              [0]
                bool bANDOR[2]
                num nSigIndex[3]
                num nSigType[3]
                num nValue[3]
            mdesc mMdesc = {leave=0}
            num nActionIndex = 60
            num nDelay = 1
            num nMoveType = 1
            num nPercentage
            num nSigValue = 1
        pointRx pPointRx[2] = {x=-395.706047, y=-287.692007, z=1039.200232, rx=-17.404604, ry=1.457158, rz=-89.580476, shoulder=lefty, elbow=epositive, wrist=wpositive}
        string sID
      [42]
        bool bMarked
        jointRx jJointRx = {j1=-133.481098, j2=-0.271586, j3=94.00243485, j4=-168.691358, j5=107.220034, j6=225.754693}
        pointRx pInter
        paraItem pParaItem
          [0]
            bool bSafePoint
            ifItem iIfItem
              [0]
                bool bANDOR[2]
                num nSigIndex[3]
                num nSigType[3]
                num nValue[3]
            mdesc mMdesc = {leave=0}
            num nActionIndex = 60
            num nDelay = 1
            num nMoveType = 1
            num nPercentage
            num nSigValue = 1
        pointRx pPointRx[2] = {x=-518.840166, y=-287.692002, z=1040.78481, rx=-17.404411, ry=1.457374, rz=-89.580244, shoulder=lefty, elbow=epositive, wrist=wpositive}
        string sID
      [43]
        bool bMarked
        jointRx jJointRx = {j1=-169.544974, j2=-34.564516, j3=135.652231, j4=-196.70666, j5=98.242514, j6=256.952537}
        pointRx pInter
        paraItem pParaItem
          [0]
            bool bSafePoint
            ifItem iIfItem
              [0]
                bool bANDOR[2]
                num nSigIndex[3]
                num nSigType[3]
                num nValue[3]
            mdesc mMdesc = {leave=0}
            num nActionIndex = 60
            num nDelay = 1
            num nMoveType = 1
            num nPercentage
            num nSigValue = 1
        pointRx pPointRx[2] = {x=-445.474256, y=-277.981159, z=882.163294, rx=16.699071, ry=0.613858, rz=-89.857323, shoulder=lefty, elbow=epositive, wrist=wpositive}
        string sID
      [44]
        bool bMarked
        jointRx jJointRx = {j1=-173.644595, j2=-34.491781, j3=138.369342, j4=-179.0487487, j5=104.740151, j6=264.0179677}
        pointRx pInter
        paraItem pParaItem
          [0]
            bool bSafePoint
            ifItem iIfItem
              [0]
                bool bANDOR[2]
                num nSigIndex[3]
                num nSigType[3]
                num nValue[3]
            mdesc mMdesc = {leave=0}
            num nActionIndex = 60
            num nDelay = 1
            num nMoveType = 1
            num nPercentage
            num nSigValue = 1
        pointRx pPointRx[2] = {x=-445.474009, y=-72.78149, z=882.163195, rx=-1.0100742, ry=0.75727, rz=-89.855065, shoulder=lefty, elbow=epositive, wrist=wpositive}
        string sID
      [45]
        bool bMarked
        jointRx jJointRx = {j1=-173.148303, j2=-23.652237, j3=75.107928, j4=-176.801258, j5=42.0835047, j6=260.997576}
        pointRx pInter
        paraItem pParaItem
          [0]
            bool bSafePoint
            ifItem iIfItem
              [0]
                bool bANDOR[2]
                num nSigIndex[3]
                num nSigType[3]
                num nValue[3]
            mdesc mMdesc = {leave=0}
            num nActionIndex = 60
            num nDelay = 1
            num nMoveType = 1
            num nPercentage
            num nSigValue = 1
        pointRx pPointRx[2] = {x=-529.449417, y=-72.791758, z=1365.530984, rx=-1.0242547, ry=-9.601326, rz=-90.0381742, shoulder=lefty, elbow=epositive, wrist=wpositive}
        string sID
      [46]
        bool bMarked
        jointRx jJointRx = {j1=-173.128911, j2=-28.821505, j3=87.506028, j4=-177.167924, j5=49.302114, j6=261.505899}
        pointRx pInter
        paraItem pParaItem
          [0]
            bool bSafePoint
            ifItem iIfItem
              [0]
                bool bANDOR[2]
                num nSigIndex[3]
                num nSigType[3]
                num nValue[3]
            mdesc mMdesc = {leave=0}
            num nActionIndex = 60
            num nDelay = 1
            num nMoveType = 1
            num nPercentage
            num nSigValue = 1
        pointRx pPointRx[2] = {x=-528.694569, y=-72.791769, z=1288.736554, rx=-1.0245197, ry=-9.602488, rz=-90.0383307, shoulder=lefty, elbow=epositive, wrist=wpositive}
        string sID
      [47]
        bool bMarked
        jointRx jJointRx = {j1=-173.184962, j2=-33.03895, j3=99.35319, j4=-177.448656, j5=56.920992, j6=262.0156524}
        pointRx pInter
        paraItem pParaItem
          [0]
            bool bSafePoint
            ifItem iIfItem
              [0]
                bool bANDOR[2]
                num nSigIndex[3]
                num nSigType[3]
                num nValue[3]
            mdesc mMdesc = {leave=0}
            num nActionIndex = 60
            num nDelay = 1
            num nMoveType = 1
            num nPercentage
            num nSigValue = 1
        pointRx pPointRx[2] = {x=-530.992203, y=-72.791768, z=1204.906755, rx=-1.0244931, ry=-9.602628, rz=-90.0383327, shoulder=lefty, elbow=epositive, wrist=wpositive}
        string sID
      [48]
        bool bMarked
        jointRx jJointRx = {j1=-173.214777, j2=-33.556097, j3=101.195834, j4=-177.491533, j5=58.243883, j6=262.117409}
        pointRx pInter
        paraItem pParaItem
          [0]
            bool bSafePoint
            ifItem iIfItem
              [0]
                bool bANDOR[2]
                num nSigIndex[3]
                num nSigType[3]
                num nValue[3]
            mdesc mMdesc = {leave=0}
            num nActionIndex = 60
            num nDelay = 1
            num nMoveType = 1
            num nPercentage
            num nSigValue = 1
        pointRx pPointRx[2] = {x=-532.232127, y=-72.791764, z=1190.718603, rx=-1.0245031, ry=-9.602735, rz=-90.0383446, shoulder=lefty, elbow=epositive, wrist=wpositive}
        string sID
      [49]
        bool bMarked
        jointRx jJointRx = {j1=-170.878262, j2=-41.834096, j3=106.133743, j4=-176.932625, j5=55.0124581, j6=259.371302}
        pointRx pInter
        paraItem pParaItem
          [0]
            bool bSafePoint
            ifItem iIfItem
              [0]
                bool bANDOR[2]
                num nSigIndex[3]
                num nSigType[3]
                num nValue[3]
            mdesc mMdesc = {leave=0}
            num nActionIndex = 60
            num nDelay = 1
            num nMoveType = 1
            num nPercentage
            num nSigValue = 1
        pointRx pPointRx[2] = {x=-459.329518, y=-72.791766, z=1175.87085, rx=-1.0239536, ry=-9.601519, rz=-90.0379744, shoulder=lefty, elbow=epositive, wrist=wpositive}
        string sID
      [50]
        bool bMarked
        jointRx jJointRx = {j1=-164.543315, j2=-49.75207, j3=106.941048, j4=-175.278138, j5=48.290196, j6=251.72242}
        pointRx pInter
        paraItem pParaItem
          [0]
            bool bSafePoint
            ifItem iIfItem
              [0]
                bool bANDOR[2]
                num nSigIndex[3]
                num nSigType[3]
                num nValue[3]
            mdesc mMdesc = {leave=0}
            num nActionIndex = 60
            num nDelay = 1
            num nMoveType = 1
            num nPercentage
            num nSigValue = 1
        pointRx pPointRx[2] = {x=-370.412471, y=-72.791755, z=1185.891907, rx=-1.0250083, ry=-9.601567, rz=-90.0385188, shoulder=lefty, elbow=epositive, wrist=wpositive}
        string sID
      [51]
        bool bMarked
        jointRx jJointRx = {j1=-150.557871, j2=-54.673707, j3=107.498981, j4=-172.114394, j5=45.209263, j6=235.417403}
        pointRx pInter
        paraItem pParaItem
          [0]
            bool bSafePoint
            ifItem iIfItem
              [0]
                bool bANDOR[2]
                num nSigIndex[3]
                num nSigType[3]
                num nValue[3]
            mdesc mMdesc = {leave=0}
            num nActionIndex = 60
            num nDelay = 1
            num nMoveType = 1
            num nPercentage
            num nSigValue = 1
        pointRx pPointRx[2] = {x=-303.196932, y=-72.792593, z=1186.264191, rx=-1.0258078, ry=-9.602273, rz=-90.0389088, shoulder=lefty, elbow=epositive, wrist=wpositive}
        string sID
      [52]
        bool bMarked
        jointRx jJointRx = {j1=-131.882073, j2=-52.891623, j3=101.937702, j4=-168.698385, j5=43.916421, j6=214.126889}
        pointRx pInter
        paraItem pParaItem
          [0]
            bool bSafePoint
            ifItem iIfItem
              [0]
                bool bANDOR[2]
                num nSigIndex[3]
                num nSigType[3]
                num nValue[3]
            mdesc mMdesc = {leave=0}
            num nActionIndex = 60
            num nDelay = 1
            num nMoveType = 1
            num nPercentage
            num nSigValue = 1
        pointRx pPointRx[2] = {x=-265.0832421, y=-72.791017, z=1226.981173, rx=-1.0236731, ry=-9.600494, rz=-90.0378745, shoulder=lefty, elbow=epositive, wrist=wpositive}
        string sID
      [53]
        bool bMarked
        jointRx jJointRx = {j1=-131.398533, j2=-48.129318, j3=93.224241, j4=-167.747499, j5=40.120899, j6=212.404386}
        pointRx pInter
        paraItem pParaItem
          [0]
            bool bSafePoint
            ifItem iIfItem
              [0]
                bool bANDOR[2]
                num nSigIndex[3]
                num nSigType[3]
                num nValue[3]
            mdesc mMdesc = {leave=0}
            num nActionIndex = 60
            num nDelay = 1
            num nMoveType = 1
            num nPercentage
            num nSigValue = 1
        pointRx pPointRx[2] = {x=-264.772643, y=-73.289439, z=1286.811055, rx=-1.0241406, ry=-9.600249, rz=-90.0380209, shoulder=lefty, elbow=epositive, wrist=wpositive}
        string sID
      [54]
        bool bMarked
        jointRx jJointRx = {j1=-144.251884, j2=-41.275682, j3=81.053431, j4=-168.18939, j5=33.105922, j6=224.769818}
        pointRx pInter
        paraItem pParaItem
          [0]
            bool bSafePoint
            ifItem iIfItem
              [0]
                bool bANDOR[2]
                num nSigIndex[3]
                num nSigType[3]
                num nValue[3]
            mdesc mMdesc = {leave=0}
            num nActionIndex = 60
            num nDelay = 1
            num nMoveType = 1
            num nPercentage
            num nSigValue = 1
        pointRx pPointRx[2] = {x=-287.116175, y=-72.447413, z=1363.274189, rx=-1.0263818, ry=-9.602793, rz=-90.03917, shoulder=lefty, elbow=epositive, wrist=wpositive}
        string sID
      [55]
        bool bMarked
        jointRx jJointRx = {j1=-161.427633, j2=-38.278204, j3=80.78039, j4=-172.806947, j5=33.91818, j6=245.804058}
        pointRx pInter
        paraItem pParaItem
          [0]
            bool bSafePoint
            ifItem iIfItem
              [0]
                bool bANDOR[2]
                num nSigIndex[3]
                num nSigType[3]
                num nValue[3]
            mdesc mMdesc = {leave=0}
            num nActionIndex = 60
            num nDelay = 1
            num nMoveType = 1
            num nPercentage
            num nSigValue = 1
        pointRx pPointRx[2] = {x=-347.943507, y=-72.792955, z=1362.805912, rx=-1.0263092, ry=-9.602341, rz=-90.0391422, shoulder=lefty, elbow=epositive, wrist=wpositive}
        string sID
      [56]
        bool bMarked
        jointRx jJointRx = {j1=-168.0500363, j2=-33.981356, j3=79.762569, j4=-175.0248349, j5=36.692248, j6=254.342934}
        pointRx pInter
        paraItem pParaItem
          [0]
            bool bSafePoint
            ifItem iIfItem
              [0]
                bool bANDOR[2]
                num nSigIndex[3]
                num nSigType[3]
                num nValue[3]
            mdesc mMdesc = {leave=0}
            num nActionIndex = 60
            num nDelay = 1
            num nMoveType = 1
            num nPercentage
            num nSigValue = 1
        pointRx pPointRx[2] = {x=-408.635334, y=-72.792697, z=1362.991056, rx=-1.0264229, ry=-9.602398, rz=-90.0392148, shoulder=lefty, elbow=epositive, wrist=wpositive}
        string sID
      [57]
        bool bMarked
        jointRx jJointRx = {j1=-164.68181, j2=-42.542405, j3=92.0793318, j4=-174.620187, j5=40.657851, j6=250.918706}
        pointRx pInter
        paraItem pParaItem
          [0]
            bool bSafePoint
            ifItem iIfItem
              [0]
                bool bANDOR[2]
                num nSigIndex[3]
                num nSigType[3]
                num nValue[3]
            mdesc mMdesc = {leave=0}
            num nActionIndex = 60
            num nDelay = 1
            num nMoveType = 1
            num nPercentage
            num nSigValue = 1
        pointRx pPointRx[2] = {x=-370.383118, y=-72.449044, z=1290.129311, rx=-1.0256153, ry=-9.601833, rz=-90.0387909, shoulder=lefty, elbow=epositive, wrist=wpositive}
        string sID
      [58]
        bool bMarked
        jointRx jJointRx = {j1=-127.503441, j2=-55.600108, j3=106.828006, j4=-168.668567, j5=46.715897, j6=210.0935795}
        pointRx pInter
        paraItem pParaItem
          [0]
            bool bSafePoint
            ifItem iIfItem
              [0]
                bool bANDOR[2]
                num nSigIndex[3]
                num nSigType[3]
                num nValue[3]
            mdesc mMdesc = {leave=0}
            num nActionIndex = 60
            num nDelay = 1
            num nMoveType = 1
            num nPercentage
            num nSigValue = 1
        pointRx pPointRx[2] = {x=-258.489334, y=-72.792581, z=1191.727111, rx=-1.024045, ry=-9.600326, rz=-90.037995, shoulder=lefty, elbow=epositive, wrist=wpositive}
        string sID
      [59]
        bool bMarked
        jointRx jJointRx = {j1=-113.574948, j2=-54.801609, j3=105.785259, j4=-167.709204, j5=48.708352, j6=195.677386}
        pointRx pInter
        paraItem pParaItem
          [0]
            bool bSafePoint
            ifItem iIfItem
              [0]
                bool bANDOR[2]
                num nSigIndex[3]
                num nSigType[3]
                num nValue[3]
            mdesc mMdesc = {leave=0}
            num nActionIndex = 60
            num nDelay = 1
            num nMoveType = 1
            num nPercentage
            num nSigValue = 1
        pointRx pPointRx[2] = {x=-239.513993, y=-72.792586, z=1199.264372, rx=-1.0254298, ry=-9.602381, rz=-90.0386982, shoulder=lefty, elbow=epositive, wrist=wpositive}
        string sID
      [60]
        bool bMarked
        jointRx jJointRx = {j1=-82.821549, j2=-56.0301157, j3=111.780274, j4=-168.953854, j5=58.457299, j6=166.854911}
        pointRx pInter
        paraItem pParaItem
          [0]
            bool bSafePoint
            ifItem iIfItem
              [0]
                bool bANDOR[2]
                num nSigIndex[3]
                num nSigType[3]
                num nValue[3]
            mdesc mMdesc = {leave=0}
            num nActionIndex = 60
            num nDelay = 1
            num nMoveType = 1
            num nPercentage
            num nSigValue = 1
        pointRx pPointRx[2] = {x=-196.990438, y=-72.792703, z=1153.733477, rx=-1.0250656, ry=-9.601957, rz=-90.0385507, shoulder=lefty, elbow=epositive, wrist=wpositive}
        string sID
      [61]
        bool bMarked
        jointRx jJointRx = {j1=-43.782169, j2=-44.715884, j3=104.221439, j4=-173.608416, j5=67.295658, j6=130.959065}
        pointRx pInter
        paraItem pParaItem
          [0]
            bool bSafePoint
            ifItem iIfItem
              [0]
                bool bANDOR[2]
                num nSigIndex[3]
                num nSigType[3]
                num nValue[3]
            mdesc mMdesc = {leave=0}
            num nActionIndex = 60
            num nDelay = 1
            num nMoveType = 1
            num nPercentage
            num nSigValue = 1
        pointRx pPointRx[2] = {x=-98.98037, y=-72.792588, z=1199.212303, rx=-1.0244226, ry=-9.602777, rz=-90.0383225, shoulder=lefty, elbow=epositive, wrist=wpositive}
        string sID
      [62]
        bool bMarked
        jointRx jJointRx = {j1=-33.126092, j2=-38.0272749, j3=100.226244, j4=-175.361365, j5=70.871203, j6=121.320684}
        pointRx pInter
        paraItem pParaItem
          [0]
            bool bSafePoint
            ifItem iIfItem
              [0]
                bool bANDOR[2]
                num nSigIndex[3]
                num nSigType[3]
                num nValue[3]
            mdesc mMdesc = {leave=0}
            num nActionIndex = 60
            num nDelay = 1
            num nMoveType = 1
            num nPercentage
            num nSigValue = 1
        pointRx pPointRx[2] = {x=-39.167207, y=-72.792342, z=1215.189033, rx=-1.0241576, ry=-9.603031, rz=-90.0382398, shoulder=lefty, elbow=epositive, wrist=wpositive}
        string sID
      [63]
        bool bMarked
        jointRx jJointRx = {j1=-26.640244, j2=-32.178556, j3=97.82685, j4=-176.491719, j5=74.724644, j6=115.49475}
        pointRx pInter
        paraItem pParaItem
          [0]
            bool bSafePoint
            ifItem iIfItem
              [0]
                bool bANDOR[2]
                num nSigIndex[3]
                num nSigType[3]
                num nValue[3]
            mdesc mMdesc = {leave=0}
            num nActionIndex = 60
            num nDelay = 1
            num nMoveType = 1
            num nPercentage
            num nSigValue = 1
        pointRx pPointRx[2] = {x=19.131819, y=-72.792471, z=1214.794054, rx=-1.0248151, ry=-9.602165, rz=-90.0383352, shoulder=lefty, elbow=epositive, wrist=wpositive}
        string sID
      [64]
        bool bMarked
        jointRx jJointRx = {j1=-31.251499, j2=-36.639218, j3=99.801437, j4=-180.984741, j5=63.657853, j6=121.825213}
        pointRx pInter
        paraItem pParaItem
          [0]
            bool bSafePoint
            ifItem iIfItem
              [0]
                bool bANDOR[2]
                num nSigIndex[3]
                num nSigType[3]
                num nValue[3]
            mdesc mMdesc = {leave=0}
            num nActionIndex = 60
            num nDelay = 1
            num nMoveType = 1
            num nPercentage
            num nSigValue = 1
        pointRx pPointRx[2] = {x=73.530888, y=-72.792474, z=1249.527518, rx=-1.00980408, ry=0.037023, rz=-89.866745, shoulder=lefty, elbow=epositive, wrist=wpositive}
        string sID
      [65]
        bool bMarked
        jointRx jJointRx = {j1=-29.625602, j2=-33.490872, j3=95.102795, j4=-181.0141949, j5=62.0826287, j6=120.237051}
        pointRx pInter
        paraItem pParaItem
          [0]
            bool bSafePoint
            ifItem iIfItem
              [0]
                bool bANDOR[2]
                num nSigIndex[3]
                num nSigType[3]
                num nValue[3]
            mdesc mMdesc = {leave=0}
            num nActionIndex = 60
            num nDelay = 1
            num nMoveType = 1
            num nPercentage
            num nSigValue = 1
        pointRx pPointRx[2] = {x=89.342541, y=-73.848982, z=1278.496301, rx=-1.00984364, ry=0.0370897, rz=-89.866758, shoulder=lefty, elbow=epositive, wrist=wpositive}
        string sID
      [66]
        bool bMarked
        jointRx jJointRx = {j1=-34.730088, j2=-32.184194, j3=84.304825, j4=-181.0689022, j5=52.670645, j6=125.515286}
        pointRx pInter
        paraItem pParaItem
          [0]
            bool bSafePoint
            ifItem iIfItem
              [0]
                bool bANDOR[2]
                num nSigIndex[3]
                num nSigType[3]
                num nValue[3]
            mdesc mMdesc = {leave=0}
            num nActionIndex = 60
            num nDelay = 1
            num nMoveType = 1
            num nPercentage
            num nSigValue = 1
        pointRx pPointRx[2] = {x=47.85983, y=-72.79225, z=1360.885028, rx=-1.00911117, ry=0.03618, rz=-89.866753, shoulder=lefty, elbow=epositive, wrist=wpositive}
        string sID
      [67]
        bool bMarked
        jointRx jJointRx = {j1=-54.722054, j2=-42.787868, j3=93.663304, j4=-180.780623, j5=51.681236, j6=145.343333}
        pointRx pInter
        paraItem pParaItem
          [0]
            bool bSafePoint
            ifItem iIfItem
              [0]
                bool bANDOR[2]
                num nSigIndex[3]
                num nSigType[3]
                num nValue[3]
            mdesc mMdesc = {leave=0}
            num nActionIndex = 60
            num nDelay = 1
            num nMoveType = 1
            num nPercentage
            num nSigValue = 1
        pointRx pPointRx[2] = {x=-39.660301, y=-72.792082, z=1314.00568418, rx=-1.00941276, ry=0.0361207, rz=-89.866728, shoulder=lefty, elbow=epositive, wrist=wpositive}
        string sID
      [68]
        bool bMarked
        jointRx jJointRx = {j1=-33.267246, j2=-42.513901, j3=112.0835977, j4=-180.919284, j5=70.0957735, j6=123.716984}
        pointRx pInter
        paraItem pParaItem
          [0]
            bool bSafePoint
            ifItem iIfItem
              [0]
                bool bANDOR[2]
                num nSigIndex[3]
                num nSigType[3]
                num nValue[3]
            mdesc mMdesc = {leave=0}
            num nActionIndex = 60
            num nDelay = 1
            num nMoveType = 1
            num nPercentage
            num nSigValue = 1
        pointRx pPointRx[2] = {x=58.0412616, y=-72.792305, z=1160.55849, rx=-1.00998313, ry=0.0362909, rz=-89.866885, shoulder=lefty, elbow=epositive, wrist=wpositive}
        string sID
      [69]
        bool bMarked
        jointRx jJointRx = {j1=-5.272998, j2=-34.693666, j3=109.0300232, j4=-181.0486852, j5=74.39402, j6=95.688496}
        pointRx pInter
        paraItem pParaItem
          [0]
            bool bSafePoint
            ifItem iIfItem
              [0]
                bool bANDOR[2]
                num nSigIndex[3]
                num nSigType[3]
                num nValue[3]
            mdesc mMdesc = {leave=0}
            num nActionIndex = 60
            num nDelay = 1
            num nMoveType = 1
            num nPercentage
            num nSigValue = 1
        pointRx pPointRx[2] = {x=138.724409, y=32.893975, z=1159.616552, rx=-1.010817, ry=0.037884, rz=-89.866801, shoulder=lefty, elbow=epositive, wrist=wpositive}
        string sID
      [70]
        bool bMarked
        jointRx jJointRx = {j1=-4.750773, j2=-30.231867, j3=104.524912, j4=-181.0486754, j5=74.34201, j6=95.167129}
        pointRx pInter
        paraItem pParaItem
          [0]
            bool bSafePoint
            ifItem iIfItem
              [0]
                bool bANDOR[2]
                num nSigIndex[3]
                num nSigType[3]
                num nValue[3]
            mdesc mMdesc = {leave=0}
            num nActionIndex = 60
            num nDelay = 1
            num nMoveType = 1
            num nPercentage
            num nSigValue = 1
        pointRx pPointRx[2] = {x=171.118595, y=32.894004, z=1180.909354, rx=-1.0101343, ry=0.0373213, rz=-89.866785, shoulder=lefty, elbow=epositive, wrist=wpositive}
        string sID
      [71]
        bool bMarked
        jointRx jJointRx = {j1=-4.653989, j2=-28.883061, j3=101.93274, j4=-181.0554282, j5=73.0969745, j6=95.0941538}
        pointRx pInter
        paraItem pParaItem
          [0]
            bool bSafePoint
            ifItem iIfItem
              [0]
                bool bANDOR[2]
                num nSigIndex[3]
                num nSigType[3]
                num nValue[3]
            mdesc mMdesc = {leave=0}
            num nActionIndex = 60
            num nDelay = 1
            num nMoveType = 1
            num nPercentage
            num nSigValue = 1
        pointRx pPointRx[2] = {x=177.941891, y=32.894009, z=1198.169889, rx=-1.0101153, ry=0.0374946, rz=-89.866798, shoulder=lefty, elbow=epositive, wrist=wpositive}
        string sID
      [72]
        bool bMarked
        jointRx jJointRx = {j1=-6.324297, j2=-43.288006, j3=121.304095, j4=-181.0301689, j5=78.0921301, j6=96.670438}
        pointRx pInter
        paraItem pParaItem
          [0]
            bool bSafePoint
            ifItem iIfItem
              [0]
                bool bANDOR[2]
                num nSigIndex[3]
                num nSigType[3]
                num nValue[3]
            mdesc mMdesc = {leave=0}
            num nActionIndex = 60
            num nDelay = 1
            num nMoveType = 1
            num nPercentage
            num nSigValue = 1
        pointRx pPointRx[2] = {x=89.587288, y=32.894025, z=1078.175922, rx=-1.0100336, ry=0.0373229, rz=-89.866767, shoulder=lefty, elbow=epositive, wrist=wpositive}
        string sID
      [73]
        bool bMarked
        jointRx jJointRx = {j1=-29.152055, j2=-40.808391, j3=117.784866, j4=-180.923594, j5=77.436909, j6=119.489453}
        pointRx pInter
        paraItem pParaItem
          [0]
            bool bSafePoint
            ifItem iIfItem
              [0]
                bool bANDOR[2]
                num nSigIndex[3]
                num nSigType[3]
                num nValue[3]
            mdesc mMdesc = {leave=0}
            num nActionIndex = 60
            num nDelay = 1
            num nMoveType = 1
            num nPercentage
            num nSigValue = 1
        pointRx pPointRx[2] = {x=91.0278996, y=-72.327826, z=1102.413174, rx=-1.0107991, ry=0.0384415, rz=-89.866785, shoulder=lefty, elbow=epositive, wrist=wpositive}
        string sID
      [74]
        bool bMarked
        jointRx jJointRx = {j1=-46.246442, j2=-55.722791, j3=128.482076, j4=-180.75609, j5=73.464404, j6=136.598984}
        pointRx pInter
        paraItem pParaItem
          [0]
            bool bSafePoint
            ifItem iIfItem
              [0]
                bool bANDOR[2]
                num nSigIndex[3]
                num nSigType[3]
                num nValue[3]
            mdesc mMdesc = {leave=0}
            num nActionIndex = 60
            num nDelay = 1
            num nMoveType = 1
            num nPercentage
            num nSigValue = 1
        pointRx pPointRx[2] = {x=-11.377417, y=-72.327654, z=1044.627758, rx=-1.00957888, ry=0.0368996, rz=-89.866787, shoulder=lefty, elbow=epositive, wrist=wpositive}
        string sID
      [75]
        bool bMarked
        jointRx jJointRx = {j1=-46.605171, j2=-57.456567, j3=132.896564, j4=-180.741462, j5=76.149251, j6=136.920045}
        pointRx pInter
        paraItem pParaItem
          [0]
            bool bSafePoint
            ifItem iIfItem
              [0]
                bool bANDOR[2]
                num nSigIndex[3]
                num nSigType[3]
                num nValue[3]
            mdesc mMdesc = {leave=0}
            num nActionIndex = 60
            num nDelay = 1
            num nMoveType = 1
            num nPercentage
            num nSigValue = 1
        pointRx pPointRx[2] = {x=-12.780183, y=-72.327727, z=1007.251626, rx=-1.00913349, ry=0.0366361, rz=-89.866763, shoulder=lefty, elbow=epositive, wrist=wpositive}
        string sID
      [76]
        bool bMarked
        jointRx jJointRx = {j1=-89.621358, j2=-69.229695, j3=134.703469, j4=-180.0469888, j5=66.483825, j6=179.773264}
        pointRx pInter
        paraItem pParaItem
          [0]
            bool bSafePoint
            ifItem iIfItem
              [0]
                bool bANDOR[2]
                num nSigIndex[3]
                num nSigType[3]
                num nValue[3]
            mdesc mMdesc = {leave=0}
            num nActionIndex = 60
            num nDelay = 1
            num nMoveType = 1
            num nPercentage
            num nSigValue = 1
        pointRx pPointRx[2] = {x=-109.0716922, y=-72.327701, z=1005.63637, rx=-1.0103058, ry=0.0364108, rz=-89.866902, shoulder=lefty, elbow=epositive, wrist=wpositive}
        string sID
      [77]
        bool bMarked
        jointRx jJointRx = {j1=-90.914117, j2=-66.731574, j3=129.968741, j4=-180.0220989, j5=64.247991, j6=181.0566361}
        pointRx pInter
        paraItem pParaItem
          [0]
            bool bSafePoint
            ifItem iIfItem
              [0]
                bool bANDOR[2]
                num nSigIndex[3]
                num nSigType[3]
                num nValue[3]
            mdesc mMdesc = {leave=0}
            num nActionIndex = 60
            num nDelay = 1
            num nMoveType = 1
            num nPercentage
            num nSigValue = 1
        pointRx pPointRx[2] = {x=-110.932852, y=-72.327788, z=1045.197534, rx=-1.0103761, ry=0.036027, rz=-89.86694, shoulder=lefty, elbow=epositive, wrist=wpositive}
        string sID
      [78]
        bool bMarked
        jointRx jJointRx = {j1=-165.265342, j2=-60.757677, j3=131.961953, j4=-178.979904, j5=71.500779, j6=255.0720448}
        pointRx pInter
        paraItem pParaItem
          [0]
            bool bSafePoint
            ifItem iIfItem
              [0]
                bool bANDOR[2]
                num nSigIndex[3]
                num nSigType[3]
                num nValue[3]
            mdesc mMdesc = {leave=0}
            num nActionIndex = 60
            num nDelay = 1
            num nMoveType = 1
            num nPercentage
            num nSigValue = 1
        pointRx pPointRx[2] = {x=-276.85417, y=-72.327729, z=1021.478785, rx=-1.0102828, ry=0.0380324, rz=-89.866783, shoulder=lefty, elbow=epositive, wrist=wpositive}
        string sID
      [79]
        bool bMarked
        jointRx jJointRx = {j1=-164.616143, j2=-57.162561, j3=122.410359, j4=-178.942453, j5=65.557451, j6=254.3092}
        pointRx pInter
        paraItem pParaItem
          [0]
            bool bSafePoint
            ifItem iIfItem
              [0]
                bool bANDOR[2]
                num nSigIndex[3]
                num nSigType[3]
                num nValue[3]
            mdesc mMdesc = {leave=0}
            num nActionIndex = 60
            num nDelay = 1
            num nMoveType = 1
            num nPercentage
            num nSigValue = 1
        pointRx pPointRx[2] = {x=-271.0494375, y=-72.327623, z=1101.43455, rx=-1.00942876, ry=0.0395777, rz=-89.86639, shoulder=lefty, elbow=epositive, wrist=wpositive}
        string sID
      [80]
        bool bMarked
        jointRx jJointRx = {j1=-172.788579, j2=-40.4338, j3=117.745846, j4=-178.978794, j5=77.478204, j6=262.698795}
        pointRx pInter
        paraItem pParaItem
          [0]
            bool bSafePoint
            ifItem iIfItem
              [0]
                bool bANDOR[2]
                num nSigIndex[3]
                num nSigType[3]
                num nValue[3]
            mdesc mMdesc = {leave=0}
            num nActionIndex = 60
            num nDelay = 1
            num nMoveType = 1
            num nPercentage
            num nSigValue = 1
        pointRx pPointRx[2] = {x=-413.537595, y=-72.3276, z=1101.399258, rx=-1.00964225, ry=0.0377699, rz=-89.866591, shoulder=lefty, elbow=epositive, wrist=wpositive}
        string sID
      [81]
        bool bMarked
        jointRx jJointRx = {j1=-172.779722, j2=-42.185789, j3=126.971722, j4=-178.999359, j5=84.950647, j6=262.823367}
        pointRx pInter
        paraItem pParaItem
          [0]
            bool bSafePoint
            ifItem iIfItem
              [0]
                bool bANDOR[2]
                num nSigIndex[3]
                num nSigType[3]
                num nValue[3]
            mdesc mMdesc = {leave=0}
            num nActionIndex = 60
            num nDelay = 1
            num nMoveType = 1
            num nPercentage
            num nSigValue = 1
        pointRx pPointRx[2] = {x=-413.202685, y=-72.327626, z=1020.485589, rx=-1.00945856, ry=0.0373518, rz=-89.866521, shoulder=lefty, elbow=epositive, wrist=wpositive}
        string sID
      [82]
        bool bMarked
        jointRx jJointRx = {j1=-173.762526, j2=-36.52442, j3=124.583138, j4=-179.000080004, j5=88.205675, j6=263.86306}
        pointRx pInter
        paraItem pParaItem
          [0]
            bool bSafePoint
            ifItem iIfItem
              [0]
                bool bANDOR[2]
                num nSigIndex[3]
                num nSigType[3]
                num nValue[3]
            mdesc mMdesc = {leave=0}
            num nActionIndex = 60
            num nDelay = 1
            num nMoveType = 1
            num nPercentage
            num nSigValue = 1
        pointRx pPointRx[2] = {x=-454.490649, y=-72.32762, z=1020.450249, rx=-1.00944981, ry=0.0372104, rz=-89.866546, shoulder=lefty, elbow=epositive, wrist=wpositive}
        string sID
      [83]
        bool bMarked
        jointRx jJointRx = {j1=-174.828859, j2=-28.228625, j3=120.323118, j4=-178.997346, j5=92.222418, j6=264.999797}
        pointRx pInter
        paraItem pParaItem
          [0]
            bool bSafePoint
            ifItem iIfItem
              [0]
                bool bANDOR[2]
                num nSigIndex[3]
                num nSigType[3]
                num nValue[3]
            mdesc mMdesc = {leave=0}
            num nActionIndex = 60
            num nDelay = 1
            num nMoveType = 1
            num nPercentage
            num nSigValue = 1
        pointRx pPointRx[2] = {x=-516.760114, y=-72.327618, z=1020.450247, rx=-1.00938216, ry=0.0374258, rz=-89.866497, shoulder=lefty, elbow=epositive, wrist=wpositive}
        string sID
      [84]
        bool bMarked
        jointRx jJointRx = {j1=-174.476731, j2=-32.134324, j3=118.120796, j4=-178.996631, j5=86.123255, j6=264.540883}
        pointRx pInter
        paraItem pParaItem
          [0]
            bool bSafePoint
            ifItem iIfItem
              [0]
                bool bANDOR[2]
                num nSigIndex[3]
                num nSigType[3]
                num nValue[3]
            mdesc mMdesc = {leave=0}
            num nActionIndex = 60
            num nDelay = 1
            num nMoveType = 1
            num nPercentage
            num nSigValue = 1
        pointRx pPointRx[2] = {x=-485.930163, y=-71.589713, z=1061.920025, rx=-1.00953266, ry=0.0391886, rz=-89.866468, shoulder=lefty, elbow=epositive, wrist=wpositive}
        string sID
      [85]
        bool bMarked
        jointRx jJointRx = {j1=-175.249335, j2=-37.428562, j3=140.970693, j4=-180.670775, j5=122.873928, j6=265.28583}
        pointRx pInter
        paraItem pParaItem
          [0]
            bool bSafePoint
            ifItem iIfItem
              [0]
                bool bANDOR[2]
                num nSigIndex[3]
                num nSigType[3]
                num nValue[3]
            mdesc mMdesc = {leave=0}
            num nActionIndex = 60
            num nDelay = 1
            num nMoveType
            num nPercentage
            num nSigValue = 1
        pointRx pPointRx[2] = {x=-228.270813, y=-62.885327, z=887.335374, rx=-1.0697583, ry=19.313004, rz=-89.513337, shoulder=lefty, elbow=epositive, wrist=wpositive}
        string sID
      [86]
        bool bMarked
        jointRx jJointRx = {j1=-55.114135, j2=-37.428562, j3=140.970693, j4=-194.186775, j5=122.873928, j6=139.07124}
        pointRx pInter
        paraItem pParaItem
          [0]
            bool bSafePoint
            ifItem iIfItem
              [0]
                bool bANDOR[2]
                num nSigIndex[3]
                num nSigType[3]
                num nValue[3]
            mdesc mMdesc = {leave=0}
            num nActionIndex = 60
            num nDelay = 1
            num nMoveType
            num nPercentage
            num nSigValue = 1
        pointRx pPointRx[2] = {x=27.333938, y=34.862636, z=815.287611, rx=-23.222857, ry=-1.370552, rz=-90.628967, shoulder=lefty, elbow=epositive, wrist=wpositive}
        string sID
      [87]
        bool bMarked
        jointRx jJointRx = {j1=13.421878, j2=-4.818376, j3=127.477265, j4=-178.119237, j5=122.0948701, j6=-9.80116}
        pointRx pInter
        paraItem pParaItem
          [0]
            bool bSafePoint
            ifItem iIfItem
              [0]
                bool bANDOR[2]
                num nSigIndex[3]
                num nSigType[3]
                num nValue[3]
            mdesc mMdesc = {leave=0}
            num nActionIndex = 60
            num nDelay = 1
            num nMoveType = 1
            num nPercentage
            num nSigValue = 1
        pointRx pPointRx[2] = {x=448.783781, y=302.866041, z=805.255089, rx=1.42221, ry=0.904693, rz=-177.39771, shoulder=lefty, elbow=epositive, wrist=wpositive}
        string sID
      [88]
        bool bMarked
        jointRx jJointRx = {j1=-0.746435, j2=38.656305, j3=103.0621354, j4=-179.633633, j5=123.453008, j6=8.386286}
        pointRx pInter
        paraItem pParaItem
          [0]
            bool bSafePoint
            ifItem iIfItem
              [0]
                bool bANDOR[2]
                num nSigIndex[3]
                num nSigType[3]
                num nValue[3]
            mdesc mMdesc = {leave=0}
            num nActionIndex = 60
            num nDelay = 1
            num nMoveType = 1
            num nPercentage
            num nSigValue = 1
        pointRx pPointRx[2] = {x=872.340958, y=193.819324, z=536.420305, rx=0.568193, ry=18.258826, rz=-172.70256, shoulder=lefty, elbow=epositive, wrist=wpositive}
        string sID
    string sID
  [PR01Washing001]
    num nFrameIndex
    num nMoveID
    num nToolIndex
    pointItem pPointItem[38]
      [0]
        bool bMarked
        jointRx jJointRx = {j1=14.463054, j2=126.686617, j3=-94.408556, j4=-18.307578, j5=-113.737208, j6=85.971215}
        pointRx pInter
        paraItem pParaItem
          [0]
            bool bSafePoint
            ifItem iIfItem
              [0]
                bool bANDOR[2]
                num nSigIndex[3]
                num nSigType[3]
                num nValue[3]
            mdesc mMdesc
            num nActionIndex = 41
            num nDelay = 1
            num nMoveType = 7
            num nPercentage
            num nSigValue
        pointRx pPointRx[2] = {x=278.890712, y=136.745171, z=230.948915, rx=84.337923, ry=-1.664851, rz=172.690172, shoulder=lefty, elbow=enegative, wrist=wnegative}
